  movel([0.496334, -1.374205, -2.584112, -0.754072, 1.570796, 2.067130],accel_mss,speed_ms,0,blend_radius_m)
  speed_ms = 0.05
  movel([0.496334, -1.321205, -2.558075, -0.833109, 1.570796, 2.067130],accel_mss,speed_ms,0,blend_radius_m)
  speed_ms = 0.051
  movel([0.496334, -1.311367, -2.552605, -0.848418, 1.570796, 2.067130],accel_mss,speed_ms,0,blend_radius_m)
  movel([0.393115, -1.332740, -2.538777, -0.840872, 1.570796, 1.963912],accel_mss,speed_ms,0,blend_radius_m)
  movel([0.393115, -1.362611, -2.554595, -0.795183, 1.570796, 1.963912],accel_mss,speed_ms,0,blend_radius_m)
  speed_ms = 0.017
  movel([0.393115, -1.394662, -2.569610, -0.748117, 1.570796, 1.963912],accel_mss,speed_ms,0,blend_radius_m)
  speed_ms = 0.051
  movel([0.404241, -1.368810, -2.587836, -0.755743, 1.570796, 1.975037],accel_mss,speed_ms,0,blend_radius_m)
  movel([0.405839, -1.365130, -2.590352, -0.756907, 1.570796, 1.976635],accel_mss,speed_ms,0,blend_radius_m)
  movel([0.405852, -1.365099, -2.590373, -0.756917, 1.570796, 1.976648],accel_mss,speed_ms,0,blend_radius_m)
  movel([0.406880, -1.363267, -2.591618, -0.757504, 1.570796, 1.977677],accel_mss,speed_ms,0,blend_radius_m)
  movel([0.408799, -1.360504, -2.593487, -0.758397, 1.570796, 1.979595],accel_mss,speed_ms,0,blend_radius_m)
  movel([0.410954, -1.358071, -2.595125, -0.759194, 1.570796, 1.981750],accel_mss,speed_ms,0,blend_radius_m)
  movel([0.413315, -1.355969, -2.596532, -0.759888, 1.570796, 1.984111],accel_mss,speed_ms,0,blend_radius_m)
  movel([0.415848, -1.354210, -2.597705, -0.760474, 1.570796, 1.986644],accel_mss,speed_ms,0,blend_radius_m)
  movel([0.418507, -1.352814, -2.598633, -0.760942, 1.570796, 1.989304],accel_mss,speed_ms,0,blend_radius_m)
  movel([0.421235, -1.351821, -2.599292, -0.761276, 1.570796, 1.992031],accel_mss,speed_ms,0,blend_radius_m)
  movel([0.423950, -1.351263, -2.599661, -0.761465, 1.570796, 1.994746],accel_mss,speed_ms,0,blend_radius_m)
  movel([0.426550, -1.351176, -2.599718, -0.761494, 1.570796, 1.997346],accel_mss,speed_ms,0,blend_radius_m)
  movel([0.428920, -1.351576, -2.599454, -0.761359, 1.570796, 1.999716],accel_mss,speed_ms,0,blend_radius_m)
  movel([0.430958, -1.352450, -2.598875, -0.761064, 1.570796, 2.001755],accel_mss,speed_ms,0,blend_radius_m)
  movel([0.432577, -1.353767, -2.598000, -0.760622, 1.570796, 2.003373],accel_mss,speed_ms,0,blend_radius_m)
  movel([0.433730, -1.355485, -2.596855, -0.760049, 1.570796, 2.004526],accel_mss,speed_ms,0,blend_radius_m)
  movel([0.434381, -1.357566, -2.595463, -0.759360, 1.570796, 2.005178],accel_mss,speed_ms,0,blend_radius_m)
  movel([0.434519, -1.359977, -2.593843, -0.758569, 1.570796, 2.005316],accel_mss,speed_ms,0,blend_radius_m)
  movel([0.434118, -1.362706, -2.591999, -0.757684, 1.570796, 2.004915],accel_mss,speed_ms,0,blend_radius_m)
  movel([0.433161, -1.365745, -2.589933, -0.756712, 1.570796, 2.003958],accel_mss,speed_ms,0,blend_radius_m)
  movel([0.431608, -1.369097, -2.587639, -0.755653, 1.570796, 2.002405],accel_mss,speed_ms,0,blend_radius_m)
  movel([0.430424, -1.371178, -2.586206, -0.755005, 1.570796, 2.001221],accel_mss,speed_ms,0,blend_radius_m)
  movel([0.439654, -1.371318, -2.586109, -0.754961, 1.570796, 2.010450],accel_mss,speed_ms,0,blend_radius_m)
  movel([0.436246, -1.378584, -2.581058, -0.752746, 1.570796, 2.007043],accel_mss,speed_ms,0,blend_radius_m)
  movel([0.410431, -1.378416, -2.581176, -0.752797, 1.570796, 1.981228],accel_mss,speed_ms,0,blend_radius_m)
  movel([0.413657, -1.371140, -2.586232, -0.755016, 1.570796, 1.984454],accel_mss,speed_ms,0,blend_radius_m)
  movel([0.422970, -1.371126, -2.586242, -0.755021, 1.570796, 1.993766],accel_mss,speed_ms,0,blend_radius_m)
  movel([0.424851, -1.367135, -2.588983, -0.756271, 1.570796, 1.995647],accel_mss,speed_ms,0,blend_radius_m)
  movel([0.425504, -1.365495, -2.590103, -0.756791, 1.570796, 1.996301],accel_mss,speed_ms,0,blend_radius_m)
  movel([0.425953, -1.364067, -2.591075, -0.757247, 1.570796, 1.996749],accel_mss,speed_ms,0,blend_radius_m)
  movel([0.426189, -1.362920, -2.591853, -0.757615, 1.570796, 1.996985],accel_mss,speed_ms,0,blend_radius_m)
  movel([0.426258, -1.361974, -2.592494, -0.757921, 1.570796, 1.997054],accel_mss,speed_ms,0,blend_radius_m)
  movel([0.426182, -1.361187, -2.593026, -0.758176, 1.570796, 1.996979],accel_mss,speed_ms,0,blend_radius_m)
  movel([0.425983, -1.360532, -2.593469, -0.758388, 1.570796, 1.996779],accel_mss,speed_ms,0,blend_radius_m)
  movel([0.425209, -1.359528, -2.594145, -0.758716, 1.570796, 1.996006],accel_mss,speed_ms,0,blend_radius_m)
  movel([0.423937, -1.358920, -2.594554, -0.758915, 1.570796, 1.994733],accel_mss,speed_ms,0,blend_radius_m)
  movel([0.422360, -1.358709, -2.594696, -0.758984, 1.570796, 1.993157],accel_mss,speed_ms,0,blend_radius_m)
  movel([0.421052, -1.358839, -2.594608, -0.758941, 1.570796, 1.991849],accel_mss,speed_ms,0,blend_radius_m)
  movel([0.419197, -1.359405, -2.594228, -0.758756, 1.570796, 1.989993],accel_mss,speed_ms,0,blend_radius_m)
  movel([0.417336, -1.360395, -2.593561, -0.758433, 1.570796, 1.988133],accel_mss,speed_ms,0,blend_radius_m)
  movel([0.415631, -1.361734, -2.592657, -0.757998, 1.570796, 1.986428],accel_mss,speed_ms,0,blend_radius_m)
  movel([0.414239, -1.363307, -2.591591, -0.757491, 1.570796, 1.985036],accel_mss,speed_ms,0,blend_radius_m)
  movel([0.413316, -1.364898, -2.590509, -0.756981, 1.570796, 1.984112],accel_mss,speed_ms,0,blend_radius_m)
  movel([0.402881, -1.388680, -2.573914, -0.749795, 1.570796, 1.973677],accel_mss,speed_ms,0,blend_radius_m)
  movel([0.400271, -1.389775, -2.573130, -0.749484, 1.570796, 1.971067],accel_mss,speed_ms,0,blend_radius_m)
  movel([0.397416, -1.391364, -2.571989, -0.749036, 1.570796, 1.968213],accel_mss,speed_ms,0,blend_radius_m)
  movel([0.394707, -1.393294, -2.570599, -0.748496, 1.570796, 1.965504],accel_mss,speed_ms,0,blend_radius_m)
  movel([0.393115, -1.394662, -2.569610, -0.748117, 1.570796, 1.963912],accel_mss,speed_ms,0,blend_radius_m)
  speed_ms = 0.05
  movel([0.393115, -1.342458, -2.544135, -0.825796, 1.570796, 1.963912],accel_mss,speed_ms,0,blend_radius_m)
  speed_ms = 0.051
  movel([0.393115, -1.332740, -2.538777, -0.840872, 1.570796, 1.963912],accel_mss,speed_ms,0,blend_radius_m)
  movel([0.435741, -1.287387, -2.567433, -0.857569, 1.570796, 2.006537],accel_mss,speed_ms,0,blend_radius_m)
  movel([0.435741, -1.318075, -2.583967, -0.810347, 1.570796, 2.006537],accel_mss,speed_ms,0,blend_radius_m)
  speed_ms = 0.017
  movel([0.435741, -1.351197, -2.599704, -0.761487, 1.570796, 2.006537],accel_mss,speed_ms,0,blend_radius_m)
  speed_ms = 0.051
  movel([0.437149, -1.352936, -2.598552, -0.760901, 1.570796, 2.007945],accel_mss,speed_ms,0,blend_radius_m)
  movel([0.438075, -1.355027, -2.597161, -0.760201, 1.570796, 2.008871],accel_mss,speed_ms,0,blend_radius_m)
  movel([0.438486, -1.357407, -2.595570, -0.759412, 1.570796, 2.009283],accel_mss,speed_ms,0,blend_radius_m)
  movel([0.438495, -1.358723, -2.594686, -0.758979, 1.570796, 2.009291],accel_mss,speed_ms,0,blend_radius_m)
  movel([0.462025, -1.359314, -2.594289, -0.758786, 1.570796, 2.032822],accel_mss,speed_ms,0,blend_radius_m)
  movel([0.462701, -1.359339, -2.594272, -0.758778, 1.570796, 2.033497],accel_mss,speed_ms,0,blend_radius_m)
  movel([0.464185, -1.359628, -2.594078, -0.758683, 1.570796, 2.034981],accel_mss,speed_ms,0,blend_radius_m)
  movel([0.465346, -1.360355, -2.593588, -0.758446, 1.570796, 2.036142],accel_mss,speed_ms,0,blend_radius_m)
  movel([0.466106, -1.361489, -2.592823, -0.758078, 1.570796, 2.036902],accel_mss,speed_ms,0,blend_radius_m)
  movel([0.466384, -1.362949, -2.591834, -0.757606, 1.570796, 2.037180],accel_mss,speed_ms,0,blend_radius_m)
  movel([0.466139, -1.364611, -2.590705, -0.757073, 1.570796, 2.036935],accel_mss,speed_ms,0,blend_radius_m)
  movel([0.465653, -1.365840, -2.589867, -0.756681, 1.570796, 2.036450],accel_mss,speed_ms,0,blend_radius_m)
  movel([0.464415, -1.367759, -2.588556, -0.756074, 1.570796, 2.035211],accel_mss,speed_ms,0,blend_radius_m)
  movel([0.463055, -1.369182, -2.587580, -0.755627, 1.570796, 2.033851],accel_mss,speed_ms,0,blend_radius_m)
  movel([0.461556, -1.370238, -2.586854, -0.755297, 1.570796, 2.032352],accel_mss,speed_ms,0,blend_radius_m)
  movel([0.459850, -1.371005, -2.586326, -0.755058, 1.570796, 2.030646],accel_mss,speed_ms,0,blend_radius_m)
  movel([0.457837, -1.371508, -2.585979, -0.754902, 1.570796, 2.028633],accel_mss,speed_ms,0,blend_radius_m)
  movel([0.455379, -1.371731, -2.585825, -0.754833, 1.570796, 2.026175],accel_mss,speed_ms,0,blend_radius_m)
  movel([0.452224, -1.371654, -2.585878, -0.754857, 1.570796, 2.023020],accel_mss,speed_ms,0,blend_radius_m)
  movel([0.450446, -1.371539, -2.585957, -0.754893, 1.570796, 2.021242],accel_mss,speed_ms,0,blend_radius_m)
  movel([0.454930, -1.362246, -2.592310, -0.757833, 1.570796, 2.025727],accel_mss,speed_ms,0,blend_radius_m)
  movel([0.447579, -1.362047, -2.592445, -0.757897, 1.570796, 2.018376],accel_mss,speed_ms,0,blend_radius_m)
  movel([0.435434, -1.387753, -2.574576, -0.750060, 1.570796, 2.006230],accel_mss,speed_ms,0,blend_radius_m)
  movel([0.442596, -1.387945, -2.574439, -0.750005, 1.570796, 2.013392],accel_mss,speed_ms,0,blend_radius_m)
  movel([0.446788, -1.379158, -2.580657, -0.752575, 1.570796, 2.017584],accel_mss,speed_ms,0,blend_radius_m)
  movel([0.446881, -1.378963, -2.580793, -0.752633, 1.570796, 2.017678],accel_mss,speed_ms,0,blend_radius_m)
  movel([0.446911, -1.378901, -2.580837, -0.752651, 1.570796, 2.017707],accel_mss,speed_ms,0,blend_radius_m)
  movel([0.450255, -1.379295, -2.580561, -0.752534, 1.570796, 2.021051],accel_mss,speed_ms,0,blend_radius_m)
  movel([0.453469, -1.379222, -2.580611, -0.752555, 1.570796, 2.024265],accel_mss,speed_ms,0,blend_radius_m)
  movel([0.456549, -1.378732, -2.580955, -0.752702, 1.570796, 2.027346],accel_mss,speed_ms,0,blend_radius_m)
  movel([0.459488, -1.377858, -2.581566, -0.752964, 1.570796, 2.030284],accel_mss,speed_ms,0,blend_radius_m)
  movel([0.462280, -1.376631, -2.582424, -0.753334, 1.570796, 2.033076],accel_mss,speed_ms,0,blend_radius_m)
  movel([0.464904, -1.375072, -2.583510, -0.753807, 1.570796, 2.035701],accel_mss,speed_ms,0,blend_radius_m)
  movel([0.467331, -1.373214, -2.584799, -0.754376, 1.570796, 2.038128],accel_mss,speed_ms,0,blend_radius_m)
  movel([0.469519, -1.371083, -2.586272, -0.755034, 1.570796, 2.040315],accel_mss,speed_ms,0,blend_radius_m)
  movel([0.471402, -1.368739, -2.587884, -0.755766, 1.570796, 2.042198],accel_mss,speed_ms,0,blend_radius_m)
  movel([0.472907, -1.366256, -2.589584, -0.756549, 1.570796, 2.043703],accel_mss,speed_ms,0,blend_radius_m)
  movel([0.473966, -1.363730, -2.591304, -0.757355, 1.570796, 2.044762],accel_mss,speed_ms,0,blend_radius_m)
  movel([0.474528, -1.361267, -2.592972, -0.758150, 1.570796, 2.045324],accel_mss,speed_ms,0,blend_radius_m)
  movel([0.474563, -1.358966, -2.594523, -0.758900, 1.570796, 2.045359],accel_mss,speed_ms,0,blend_radius_m)
  movel([0.474065, -1.356904, -2.595906, -0.759578, 1.570796, 2.044861],accel_mss,speed_ms,0,blend_radius_m)
  movel([0.473042, -1.355135, -2.597089, -0.760165, 1.570796, 2.043838],accel_mss,speed_ms,0,blend_radius_m)
  movel([0.471495, -1.353700, -2.598045, -0.760644, 1.570796, 2.042292],accel_mss,speed_ms,0,blend_radius_m)
  movel([0.469420, -1.352631, -2.598755, -0.761004, 1.570796, 2.040217],accel_mss,speed_ms,0,blend_radius_m)
  movel([0.466801, -1.351958, -2.599201, -0.761230, 1.570796, 2.037597],accel_mss,speed_ms,0,blend_radius_m)
  movel([0.466254, -1.351881, -2.599252, -0.761256, 1.570796, 2.037050],accel_mss,speed_ms,0,blend_radius_m)
  movel([0.435741, -1.351197, -2.599704, -0.761487, 1.570796, 2.006537],accel_mss,speed_ms,0,blend_radius_m)
  speed_ms = 0.05
  movel([0.435741, -1.297350, -2.573030, -0.842009, 1.570796, 2.006537],accel_mss,speed_ms,0,blend_radius_m)
  speed_ms = 0.051
  movel([0.435741, -1.287387, -2.567433, -0.857569, 1.570796, 2.006537],accel_mss,speed_ms,0,blend_radius_m)
  movel([0.468006, -1.313184, -2.551452, -0.847754, 1.570796, 2.038802],accel_mss,speed_ms,0,blend_radius_m)
  movel([0.468006, -1.343421, -2.567577, -0.801391, 1.570796, 2.038802],accel_mss,speed_ms,0,blend_radius_m)
  speed_ms = 0.017
  movel([0.468006, -1.375946, -2.582901, -0.753542, 1.570796, 2.038802],accel_mss,speed_ms,0,blend_radius_m)
  speed_ms = 0.051
  movel([0.456016, -1.400133, -2.565628, -0.746628, 1.570796, 2.026813],accel_mss,speed_ms,0,blend_radius_m)
  movel([0.453789, -1.404662, -2.562298, -0.745429, 1.570796, 2.024585],accel_mss,speed_ms,0,blend_radius_m)
  movel([0.453641, -1.404968, -2.562072, -0.745349, 1.570796, 2.024437],accel_mss,speed_ms,0,blend_radius_m)
  movel([0.452579, -1.406671, -2.560812, -0.744907, 1.570796, 2.023375],accel_mss,speed_ms,0,blend_radius_m)
  movel([0.450661, -1.409191, -2.558938, -0.744260, 1.570796, 2.021458],accel_mss,speed_ms,0,blend_radius_m)
  movel([0.448563, -1.411364, -2.557315, -0.743710, 1.570796, 2.019359],accel_mss,speed_ms,0,blend_radius_m)
  movel([0.446304, -1.413204, -2.555935, -0.743250, 1.570796, 2.017100],accel_mss,speed_ms,0,blend_radius_m)
  movel([0.443919, -1.414710, -2.554802, -0.742877, 1.570796, 2.014715],accel_mss,speed_ms,0,blend_radius_m)
  movel([0.441440, -1.415871, -2.553926, -0.742592, 1.570796, 2.012236],accel_mss,speed_ms,0,blend_radius_m)
  movel([0.438915, -1.416664, -2.553326, -0.742399, 1.570796, 2.009711],accel_mss,speed_ms,0,blend_radius_m)
  movel([0.436416, -1.417065, -2.553023, -0.742301, 1.570796, 2.007212],accel_mss,speed_ms,0,blend_radius_m)
  movel([0.434024, -1.417050, -2.553035, -0.742305, 1.570796, 2.004820],accel_mss,speed_ms,0,blend_radius_m)
  movel([0.431843, -1.416611, -2.553367, -0.742411, 1.570796, 2.002639],accel_mss,speed_ms,0,blend_radius_m)
  movel([0.429962, -1.415757, -2.554012, -0.742620, 1.570796, 2.000758],accel_mss,speed_ms,0,blend_radius_m)
  movel([0.428455, -1.414516, -2.554948, -0.742925, 1.570796, 1.999251],accel_mss,speed_ms,0,blend_radius_m)
  movel([0.427374, -1.412916, -2.556151, -0.743322, 1.570796, 1.998171],accel_mss,speed_ms,0,blend_radius_m)
  movel([0.426747, -1.410989, -2.557595, -0.743804, 1.570796, 1.997543],accel_mss,speed_ms,0,blend_radius_m)
  movel([0.426600, -1.408754, -2.559264, -0.744372, 1.570796, 1.997396],accel_mss,speed_ms,0,blend_radius_m)
  movel([0.426957, -1.406212, -2.561152, -0.745025, 1.570796, 1.997753],accel_mss,speed_ms,0,blend_radius_m)
  movel([0.427853, -1.403363, -2.563256, -0.745769, 1.570796, 1.998650],accel_mss,speed_ms,0,blend_radius_m)
  movel([0.429335, -1.400194, -2.565584, -0.746612, 1.570796, 2.000131],accel_mss,speed_ms,0,blend_radius_m)
  movel([0.430468, -1.398225, -2.567022, -0.747142, 1.570796, 2.001264],accel_mss,speed_ms,0,blend_radius_m)
  movel([0.421486, -1.398069, -2.567136, -0.747184, 1.570796, 1.992282],accel_mss,speed_ms,0,blend_radius_m)
  movel([0.424715, -1.391019, -2.572237, -0.749133, 1.570796, 1.995511],accel_mss,speed_ms,0,blend_radius_m)
  movel([0.449964, -1.391682, -2.571760, -0.748946, 1.570796, 2.020760],accel_mss,speed_ms,0,blend_radius_m)
  movel([0.446570, -1.398709, -2.566669, -0.747011, 1.570796, 2.017367],accel_mss,speed_ms,0,blend_radius_m)
  movel([0.437657, -1.398406, -2.566890, -0.747093, 1.570796, 2.008453],accel_mss,speed_ms,0,blend_radius_m)
  movel([0.435797, -1.402197, -2.564115, -0.746078, 1.570796, 2.006593],accel_mss,speed_ms,0,blend_radius_m)
  movel([0.435154, -1.403745, -2.562975, -0.745669, 1.570796, 2.005951],accel_mss,speed_ms,0,blend_radius_m)
  movel([0.434713, -1.405089, -2.561983, -0.745317, 1.570796, 2.005509],accel_mss,speed_ms,0,blend_radius_m)
  movel([0.434481, -1.406166, -2.561185, -0.745037, 1.570796, 2.005277],accel_mss,speed_ms,0,blend_radius_m)
  movel([0.434406, -1.407058, -2.560524, -0.744807, 1.570796, 2.005202],accel_mss,speed_ms,0,blend_radius_m)
  movel([0.434470, -1.407800, -2.559974, -0.744616, 1.570796, 2.005266],accel_mss,speed_ms,0,blend_radius_m)
  movel([0.434651, -1.408420, -2.559512, -0.744457, 1.570796, 2.005447],accel_mss,speed_ms,0,blend_radius_m)
  movel([0.435365, -1.409380, -2.558797, -0.744212, 1.570796, 2.006161],accel_mss,speed_ms,0,blend_radius_m)
  movel([0.436549, -1.409986, -2.558345, -0.744058, 1.570796, 2.007345],accel_mss,speed_ms,0,blend_radius_m)
  movel([0.438023, -1.410235, -2.558159, -0.743995, 1.570796, 2.008819],accel_mss,speed_ms,0,blend_radius_m)
  movel([0.439241, -1.410163, -2.558213, -0.744013, 1.570796, 2.010038],accel_mss,speed_ms,0,blend_radius_m)
  movel([0.440983, -1.409705, -2.558554, -0.744129, 1.570796, 2.011779],accel_mss,speed_ms,0,blend_radius_m)
  movel([0.442739, -1.408855, -2.559189, -0.744346, 1.570796, 2.013535],accel_mss,speed_ms,0,blend_radius_m)
  movel([0.444367, -1.407667, -2.560072, -0.744650, 1.570796, 2.015163],accel_mss,speed_ms,0,blend_radius_m)
  movel([0.445716, -1.406238, -2.561132, -0.745018, 1.570796, 2.016512],accel_mss,speed_ms,0,blend_radius_m)
  movel([0.446637, -1.404764, -2.562223, -0.745402, 1.570796, 2.017433],accel_mss,speed_ms,0,blend_radius_m)
  movel([0.457925, -1.381620, -2.578926, -0.751843, 1.570796, 2.028721],accel_mss,speed_ms,0,blend_radius_m)
  movel([0.460558, -1.380630, -2.579623, -0.752136, 1.570796, 2.031354],accel_mss,speed_ms,0,blend_radius_m)
  movel([0.463484, -1.379143, -2.580667, -0.752579, 1.570796, 2.034281],accel_mss,speed_ms,0,blend_radius_m)
  movel([0.466307, -1.377290, -2.581964, -0.753135, 1.570796, 2.037103],accel_mss,speed_ms,0,blend_radius_m)
  movel([0.468006, -1.375946, -2.582901, -0.753542, 1.570796, 2.038802],accel_mss,speed_ms,0,blend_radius_m)
  speed_ms = 0.05
  movel([0.468006, -1.323012, -2.556913, -0.832464, 1.570796, 2.038802],accel_mss,speed_ms,0,blend_radius_m)
  speed_ms = 0.051
  movel([0.468006, -1.313184, -2.551452, -0.847754, 1.570796, 2.038802],accel_mss,speed_ms,0,blend_radius_m)
  movel([0.425547, -1.355903, -2.523122, -0.833364, 1.570796, 1.996343],accel_mss,speed_ms,0,blend_radius_m)
  movel([0.425547, -1.385315, -2.538580, -0.788493, 1.570796, 1.996343],accel_mss,speed_ms,0,blend_radius_m)
  speed_ms = 0.017
  movel([0.425547, -1.416785, -2.553235, -0.742369, 1.570796, 1.996343],accel_mss,speed_ms,0,blend_radius_m)
  speed_ms = 0.051
  movel([0.403473, -1.416474, -2.553470, -0.742445, 1.570796, 1.974270],accel_mss,speed_ms,0,blend_radius_m)
  movel([0.396842, -1.416472, -2.553471, -0.742445, 1.570796, 1.967639],accel_mss,speed_ms,0,blend_radius_m)
  movel([0.396831, -1.416472, -2.553471, -0.742445, 1.570796, 1.967627],accel_mss,speed_ms,0,blend_radius_m)
  movel([0.395180, -1.416267, -2.553626, -0.742495, 1.570796, 1.965977],accel_mss,speed_ms,0,blend_radius_m)
  movel([0.392846, -1.415632, -2.554106, -0.742651, 1.570796, 1.963642],accel_mss,speed_ms,0,blend_radius_m)
  movel([0.390981, -1.414656, -2.554843, -0.742891, 1.570796, 1.961777],accel_mss,speed_ms,0,blend_radius_m)
  movel([0.389571, -1.413365, -2.555814, -0.743210, 1.570796, 1.960368],accel_mss,speed_ms,0,blend_radius_m)
  movel([0.388609, -1.411785, -2.557000, -0.743604, 1.570796, 1.959406],accel_mss,speed_ms,0,blend_radius_m)
  movel([0.388105, -1.409938, -2.558381, -0.744070, 1.570796, 1.958902],accel_mss,speed_ms,0,blend_radius_m)
  movel([0.388072, -1.407859, -2.559929, -0.744600, 1.570796, 1.958868],accel_mss,speed_ms,0,blend_radius_m)
  movel([0.388518, -1.405604, -2.561602, -0.745183, 1.570796, 1.959314],accel_mss,speed_ms,0,blend_radius_m)
  movel([0.389446, -1.403245, -2.563343, -0.745801, 1.570796, 1.960243],accel_mss,speed_ms,0,blend_radius_m)
  movel([0.390831, -1.400879, -2.565081, -0.746428, 1.570796, 1.961628],accel_mss,speed_ms,0,blend_radius_m)
  movel([0.392628, -1.398602, -2.566747, -0.747040, 1.570796, 1.963425],accel_mss,speed_ms,0,blend_radius_m)
  movel([0.394772, -1.396508, -2.568271, -0.747609, 1.570796, 1.965569],accel_mss,speed_ms,0,blend_radius_m)
  movel([0.397198, -1.394665, -2.569608, -0.748116, 1.570796, 1.967995],accel_mss,speed_ms,0,blend_radius_m)
  movel([0.399853, -1.393125, -2.570721, -0.748543, 1.570796, 1.970650],accel_mss,speed_ms,0,blend_radius_m)
  movel([0.402697, -1.391919, -2.571590, -0.748880, 1.570796, 1.973493],accel_mss,speed_ms,0,blend_radius_m)
  movel([0.405704, -1.391081, -2.572193, -0.749115, 1.570796, 1.976501],accel_mss,speed_ms,0,blend_radius_m)
  movel([0.408860, -1.390644, -2.572506, -0.749238, 1.570796, 1.979657],accel_mss,speed_ms,0,blend_radius_m)
  movel([0.412150, -1.390646, -2.572505, -0.749238, 1.570796, 1.982946],accel_mss,speed_ms,0,blend_radius_m)
  movel([0.414108, -1.390866, -2.572347, -0.749176, 1.570796, 1.984905],accel_mss,speed_ms,0,blend_radius_m)
  movel([0.418149, -1.381867, -2.578751, -0.751770, 1.570796, 1.988945],accel_mss,speed_ms,0,blend_radius_m)
  movel([0.425423, -1.381914, -2.578718, -0.751757, 1.570796, 1.996219],accel_mss,speed_ms,0,blend_radius_m)
  movel([0.414112, -1.406828, -2.560695, -0.744866, 1.570796, 1.984908],accel_mss,speed_ms,0,blend_radius_m)
  movel([0.407010, -1.406787, -2.560726, -0.744877, 1.570796, 1.977806],accel_mss,speed_ms,0,blend_radius_m)
  movel([0.410920, -1.398011, -2.567178, -0.747200, 1.570796, 1.981717],accel_mss,speed_ms,0,blend_radius_m)
  movel([0.407049, -1.397939, -2.567230, -0.747220, 1.570796, 1.977845],accel_mss,speed_ms,0,blend_radius_m)
  movel([0.405413, -1.398026, -2.567167, -0.747196, 1.570796, 1.976209],accel_mss,speed_ms,0,blend_radius_m)
  movel([0.403942, -1.398220, -2.567026, -0.747143, 1.570796, 1.974739],accel_mss,speed_ms,0,blend_radius_m)
  movel([0.402713, -1.398494, -2.566826, -0.747069, 1.570796, 1.973509],accel_mss,speed_ms,0,blend_radius_m)
  movel([0.401648, -1.398841, -2.566572, -0.746975, 1.570796, 1.972444],accel_mss,speed_ms,0,blend_radius_m)
  movel([0.400712, -1.399250, -2.566274, -0.746865, 1.570796, 1.971508],accel_mss,speed_ms,0,blend_radius_m)
  movel([0.399874, -1.399720, -2.565930, -0.746739, 1.570796, 1.970671],accel_mss,speed_ms,0,blend_radius_m)
  movel([0.398410, -1.400878, -2.565082, -0.746428, 1.570796, 1.969206],accel_mss,speed_ms,0,blend_radius_m)
  movel([0.397202, -1.402325, -2.564020, -0.746044, 1.570796, 1.967999],accel_mss,speed_ms,0,blend_radius_m)
  movel([0.396320, -1.403889, -2.562869, -0.745631, 1.570796, 1.967117],accel_mss,speed_ms,0,blend_radius_m)
  movel([0.395938, -1.405045, -2.562015, -0.745329, 1.570796, 1.966735],accel_mss,speed_ms,0,blend_radius_m)
  movel([0.395831, -1.406526, -2.560919, -0.744944, 1.570796, 1.966627],accel_mss,speed_ms,0,blend_radius_m)
  movel([0.396199, -1.407832, -2.559950, -0.744608, 1.570796, 1.966995],accel_mss,speed_ms,0,blend_radius_m)
  movel([0.397028, -1.408849, -2.559193, -0.744347, 1.570796, 1.967824],accel_mss,speed_ms,0,blend_radius_m)
  movel([0.398251, -1.409481, -2.558722, -0.744186, 1.570796, 1.969048],accel_mss,speed_ms,0,blend_radius_m)
  movel([0.399687, -1.409681, -2.558573, -0.744135, 1.570796, 1.970483],accel_mss,speed_ms,0,blend_radius_m)
  movel([0.422863, -1.409863, -2.558437, -0.744089, 1.570796, 1.993659],accel_mss,speed_ms,0,blend_radius_m)
  movel([0.422993, -1.411906, -2.556909, -0.743574, 1.570796, 1.993789],accel_mss,speed_ms,0,blend_radius_m)
  movel([0.423592, -1.413991, -2.555343, -0.743055, 1.570796, 1.994388],accel_mss,speed_ms,0,blend_radius_m)
  movel([0.424651, -1.415802, -2.553978, -0.742609, 1.570796, 1.995448],accel_mss,speed_ms,0,blend_radius_m)
  movel([0.425547, -1.416785, -2.553235, -0.742369, 1.570796, 1.996343],accel_mss,speed_ms,0,blend_radius_m)
  speed_ms = 0.05
  movel([0.425547, -1.365481, -2.528361, -0.818547, 1.570796, 1.996343],accel_mss,speed_ms,0,blend_radius_m)
  speed_ms = 0.051
  movel([0.425547, -1.355903, -2.523122, -0.833364, 1.570796, 1.996343],accel_mss,speed_ms,0,blend_radius_m)
  movel([0.496386, -1.351291, -2.526295, -0.834803, 1.570796, 2.067183],accel_mss,speed_ms,0,blend_radius_m)
  movel([0.496386, -1.380797, -2.541825, -0.789767, 1.570796, 2.067183],accel_mss,speed_ms,0,blend_radius_m)
  speed_ms = 0.017
  movel([0.496386, -1.412384, -2.556551, -0.743454, 1.570796, 2.067183],accel_mss,speed_ms,0,blend_radius_m)
  speed_ms = 0.051
  movel([0.494250, -1.412916, -2.556152, -0.743322, 1.570796, 2.065047],accel_mss,speed_ms,0,blend_radius_m)
  movel([0.492155, -1.413824, -2.555469, -0.743096, 1.570796, 2.062951],accel_mss,speed_ms,0,blend_radius_m)
  movel([0.490635, -1.414706, -2.554805, -0.742878, 1.570796, 2.061431],accel_mss,speed_ms,0,blend_radius_m)
  movel([0.498563, -1.433670, -2.540242, -0.738476, 1.570796, 2.069360],accel_mss,speed_ms,0,blend_radius_m)
  movel([0.507323, -1.428619, -2.544174, -0.739595, 1.570796, 2.078119],accel_mss,speed_ms,0,blend_radius_m)
  movel([0.504979, -1.429334, -2.543621, -0.739435, 1.570796, 2.075776],accel_mss,speed_ms,0,blend_radius_m)
  movel([0.502994, -1.429562, -2.543443, -0.739383, 1.570796, 2.073791],accel_mss,speed_ms,0,blend_radius_m)
  movel([0.501213, -1.429380, -2.543585, -0.739424, 1.570796, 2.072009],accel_mss,speed_ms,0,blend_radius_m)
  movel([0.499589, -1.428783, -2.544047, -0.739558, 1.570796, 2.070385],accel_mss,speed_ms,0,blend_radius_m)
  movel([0.498113, -1.427739, -2.544855, -0.739794, 1.570796, 2.068909],accel_mss,speed_ms,0,blend_radius_m)
  movel([0.496789, -1.426184, -2.546056, -0.740149, 1.570796, 2.067585],accel_mss,speed_ms,0,blend_radius_m)
  movel([0.495653, -1.424054, -2.547695, -0.740640, 1.570796, 2.066450],accel_mss,speed_ms,0,blend_radius_m)
  movel([0.495357, -1.423295, -2.548277, -0.740817, 1.570796, 2.066154],accel_mss,speed_ms,0,blend_radius_m)
  movel([0.496802, -1.422585, -2.548821, -0.740983, 1.570796, 2.067599],accel_mss,speed_ms,0,blend_radius_m)
  movel([0.498935, -1.421858, -2.549377, -0.741154, 1.570796, 2.069732],accel_mss,speed_ms,0,blend_radius_m)
  movel([0.501190, -1.421465, -2.549677, -0.741247, 1.570796, 2.071986],accel_mss,speed_ms,0,blend_radius_m)
  movel([0.503721, -1.421404, -2.549724, -0.741261, 1.570796, 2.074517],accel_mss,speed_ms,0,blend_radius_m)
  movel([0.506892, -1.421700, -2.549497, -0.741191, 1.570796, 2.077688],accel_mss,speed_ms,0,blend_radius_m)
  movel([0.508953, -1.421976, -2.549287, -0.741126, 1.570796, 2.079749],accel_mss,speed_ms,0,blend_radius_m)
  movel([0.511017, -1.422212, -2.549106, -0.741071, 1.570796, 2.081813],accel_mss,speed_ms,0,blend_radius_m)
  movel([0.512879, -1.422311, -2.549031, -0.741048, 1.570796, 2.083675],accel_mss,speed_ms,0,blend_radius_m)
  movel([0.514361, -1.422273, -2.549060, -0.741057, 1.570796, 2.085157],accel_mss,speed_ms,0,blend_radius_m)
  movel([0.516717, -1.421930, -2.549322, -0.741137, 1.570796, 2.087514],accel_mss,speed_ms,0,blend_radius_m)
  movel([0.519106, -1.421259, -2.549835, -0.741296, 1.570796, 2.089902],accel_mss,speed_ms,0,blend_radius_m)
  movel([0.521253, -1.420298, -2.550567, -0.741524, 1.570796, 2.092049],accel_mss,speed_ms,0,blend_radius_m)
  movel([0.523071, -1.419109, -2.551472, -0.741808, 1.570796, 2.093867],accel_mss,speed_ms,0,blend_radius_m)
  movel([0.524605, -1.417699, -2.552542, -0.742147, 1.570796, 2.095402],accel_mss,speed_ms,0,blend_radius_m)
  movel([0.525885, -1.416058, -2.553785, -0.742546, 1.570796, 2.096681],accel_mss,speed_ms,0,blend_radius_m)
  movel([0.526903, -1.414161, -2.555215, -0.743013, 1.570796, 2.097699],accel_mss,speed_ms,0,blend_radius_m)
  movel([0.527617, -1.412010, -2.556831, -0.743548, 1.570796, 2.098413],accel_mss,speed_ms,0,blend_radius_m)
  movel([0.527962, -1.409636, -2.558606, -0.744147, 1.570796, 2.098758],accel_mss,speed_ms,0,blend_radius_m)
  movel([0.527865, -1.407145, -2.560460, -0.744784, 1.570796, 2.098662],accel_mss,speed_ms,0,blend_radius_m)
  movel([0.527282, -1.404723, -2.562253, -0.745413, 1.570796, 2.098079],accel_mss,speed_ms,0,blend_radius_m)
  movel([0.526229, -1.402597, -2.563820, -0.745972, 1.570796, 2.097026],accel_mss,speed_ms,0,blend_radius_m)
  movel([0.524809, -1.400967, -2.565017, -0.746405, 1.570796, 2.095605],accel_mss,speed_ms,0,blend_radius_m)
  movel([0.523535, -1.400104, -2.565650, -0.746636, 1.570796, 2.094332],accel_mss,speed_ms,0,blend_radius_m)
  movel([0.522574, -1.399712, -2.565936, -0.746741, 1.570796, 2.093370],accel_mss,speed_ms,0,blend_radius_m)
  movel([0.521144, -1.399562, -2.566046, -0.746781, 1.570796, 2.091941],accel_mss,speed_ms,0,blend_radius_m)
  movel([0.519713, -1.399841, -2.565842, -0.746706, 1.570796, 2.090509],accel_mss,speed_ms,0,blend_radius_m)
  movel([0.518321, -1.400499, -2.565360, -0.746530, 1.570796, 2.089117],accel_mss,speed_ms,0,blend_radius_m)
  movel([0.517042, -1.401495, -2.564630, -0.746264, 1.570796, 2.087839],accel_mss,speed_ms,0,blend_radius_m)
  movel([0.516004, -1.402743, -2.563713, -0.745933, 1.570796, 2.086801],accel_mss,speed_ms,0,blend_radius_m)
  movel([0.515361, -1.404091, -2.562720, -0.745578, 1.570796, 2.086157],accel_mss,speed_ms,0,blend_radius_m)
  movel([0.515210, -1.405299, -2.561828, -0.745262, 1.570796, 2.086007],accel_mss,speed_ms,0,blend_radius_m)
  movel([0.515554, -1.406380, -2.561027, -0.744982, 1.570796, 2.086350],accel_mss,speed_ms,0,blend_radius_m)
  movel([0.516416, -1.407204, -2.560416, -0.744769, 1.570796, 2.087212],accel_mss,speed_ms,0,blend_radius_m)
  movel([0.517279, -1.407592, -2.560128, -0.744669, 1.570796, 2.088075],accel_mss,speed_ms,0,blend_radius_m)
  movel([0.518096, -1.407710, -2.560040, -0.744639, 1.570796, 2.088893],accel_mss,speed_ms,0,blend_radius_m)
  movel([0.519202, -1.407488, -2.560205, -0.744696, 1.570796, 2.089998],accel_mss,speed_ms,0,blend_radius_m)
  movel([0.520433, -1.406863, -2.560669, -0.744857, 1.570796, 2.091230],accel_mss,speed_ms,0,blend_radius_m)
  movel([0.521857, -1.405770, -2.561479, -0.745140, 1.570796, 2.092653],accel_mss,speed_ms,0,blend_radius_m)
  movel([0.523464, -1.404168, -2.562663, -0.745558, 1.570796, 2.094260],accel_mss,speed_ms,0,blend_radius_m)
  movel([0.523573, -1.404048, -2.562751, -0.745589, 1.570796, 2.094369],accel_mss,speed_ms,0,blend_radius_m)
  movel([0.524385, -1.403902, -2.562859, -0.745628, 1.570796, 2.095181],accel_mss,speed_ms,0,blend_radius_m)
  movel([0.525389, -1.404028, -2.562766, -0.745595, 1.570796, 2.096185],accel_mss,speed_ms,0,blend_radius_m)
  movel([0.526064, -1.404552, -2.562380, -0.745458, 1.570796, 2.096860],accel_mss,speed_ms,0,blend_radius_m)
  movel([0.526402, -1.405475, -2.561697, -0.745217, 1.570796, 2.097199],accel_mss,speed_ms,0,blend_radius_m)
  movel([0.526323, -1.406784, -2.560727, -0.744877, 1.570796, 2.097119],accel_mss,speed_ms,0,blend_radius_m)
  movel([0.525762, -1.408332, -2.559577, -0.744479, 1.570796, 2.096558],accel_mss,speed_ms,0,blend_radius_m)
  movel([0.524768, -1.409827, -2.558464, -0.744098, 1.570796, 2.095564],accel_mss,speed_ms,0,blend_radius_m)
  movel([0.524179, -1.410451, -2.557998, -0.743940, 1.570796, 2.094975],accel_mss,speed_ms,0,blend_radius_m)
  movel([0.523546, -1.410986, -2.557598, -0.743805, 1.570796, 2.094342],accel_mss,speed_ms,0,blend_radius_m)
  movel([0.522160, -1.411793, -2.556994, -0.743602, 1.570796, 2.092957],accel_mss,speed_ms,0,blend_radius_m)
  movel([0.522122, -1.411809, -2.556982, -0.743598, 1.570796, 2.092918],accel_mss,speed_ms,0,blend_radius_m)
  movel([0.520402, -1.412510, -2.556456, -0.743423, 1.570796, 2.091198],accel_mss,speed_ms,0,blend_radius_m)
  movel([0.518013, -1.413155, -2.555972, -0.743262, 1.570796, 2.088809],accel_mss,speed_ms,0,blend_radius_m)
  movel([0.515460, -1.413467, -2.555737, -0.743185, 1.570796, 2.086257],accel_mss,speed_ms,0,blend_radius_m)
  movel([0.512586, -1.413441, -2.555757, -0.743191, 1.570796, 2.083382],accel_mss,speed_ms,0,blend_radius_m)
  movel([0.509044, -1.413037, -2.556060, -0.743292, 1.570796, 2.079841],accel_mss,speed_ms,0,blend_radius_m)
  movel([0.506535, -1.412642, -2.556357, -0.743390, 1.570796, 2.077331],accel_mss,speed_ms,0,blend_radius_m)
  movel([0.504024, -1.412280, -2.556629, -0.743481, 1.570796, 2.074820],accel_mss,speed_ms,0,blend_radius_m)
  movel([0.501612, -1.412053, -2.556799, -0.743537, 1.570796, 2.072409],accel_mss,speed_ms,0,blend_radius_m)
  movel([0.499823, -1.412015, -2.556827, -0.743547, 1.570796, 2.070619],accel_mss,speed_ms,0,blend_radius_m)
  movel([0.498273, -1.412102, -2.556762, -0.743525, 1.570796, 2.069069],accel_mss,speed_ms,0,blend_radius_m)
  movel([0.496386, -1.412384, -2.556551, -0.743454, 1.570796, 2.067183],accel_mss,speed_ms,0,blend_radius_m)
  speed_ms = 0.05
  movel([0.496386, -1.360898, -2.531558, -0.819933, 1.570796, 2.067183],accel_mss,speed_ms,0,blend_radius_m)
  speed_ms = 0.051
  movel([0.496386, -1.351291, -2.526295, -0.834803, 1.570796, 2.067183],accel_mss,speed_ms,0,blend_radius_m)
  movel([0.501294, -1.380106, -2.506003, -0.826280, 1.570796, 2.072091],accel_mss,speed_ms,0,blend_radius_m)
  movel([0.501294, -1.409013, -2.521091, -0.782286, 1.570796, 2.072091],accel_mss,speed_ms,0,blend_radius_m)
  speed_ms = 0.017
  movel([0.501294, -1.439855, -2.535375, -0.737159, 1.570796, 2.072091],accel_mss,speed_ms,0,blend_radius_m)
  speed_ms = 0.051
  movel([0.501364, -1.438344, -2.536570, -0.737475, 1.570796, 2.072160],accel_mss,speed_ms,0,blend_radius_m)
  movel([0.501902, -1.436575, -2.537964, -0.737850, 1.570796, 2.072698],accel_mss,speed_ms,0,blend_radius_m)
  movel([0.502852, -1.434869, -2.539304, -0.738216, 1.570796, 2.073649],accel_mss,speed_ms,0,blend_radius_m)
  movel([0.503411, -1.434165, -2.539855, -0.738369, 1.570796, 2.074207],accel_mss,speed_ms,0,blend_radius_m)
  movel([0.503999, -1.433568, -2.540323, -0.738498, 1.570796, 2.074796],accel_mss,speed_ms,0,blend_radius_m)
  movel([0.504606, -1.433084, -2.540701, -0.738604, 1.570796, 2.075402],accel_mss,speed_ms,0,blend_radius_m)
  movel([0.505876, -1.432412, -2.541226, -0.738751, 1.570796, 2.076673],accel_mss,speed_ms,0,blend_radius_m)
  movel([0.507182, -1.432148, -2.541432, -0.738809, 1.570796, 2.077978],accel_mss,speed_ms,0,blend_radius_m)
  movel([0.508066, -1.432194, -2.541395, -0.738799, 1.570796, 2.078863],accel_mss,speed_ms,0,blend_radius_m)
  movel([0.509244, -1.432844, -2.540888, -0.738657, 1.570796, 2.080041],accel_mss,speed_ms,0,blend_radius_m)
  movel([0.509920, -1.433743, -2.540185, -0.738460, 1.570796, 2.080716],accel_mss,speed_ms,0,blend_radius_m)
  movel([0.510117, -1.434828, -2.539336, -0.738225, 1.570796, 2.080914],accel_mss,speed_ms,0,blend_radius_m)
  movel([0.509853, -1.436017, -2.538403, -0.737969, 1.570796, 2.080649],accel_mss,speed_ms,0,blend_radius_m)
  movel([0.509157, -1.437210, -2.537464, -0.737715, 1.570796, 2.079953],accel_mss,speed_ms,0,blend_radius_m)
  movel([0.508088, -1.438286, -2.536615, -0.737487, 1.570796, 2.078884],accel_mss,speed_ms,0,blend_radius_m)
  movel([0.506729, -1.439143, -2.535939, -0.737307, 1.570796, 2.077525],accel_mss,speed_ms,0,blend_radius_m)
  movel([0.505151, -1.439703, -2.535495, -0.737190, 1.570796, 2.075947],accel_mss,speed_ms,0,blend_radius_m)
  movel([0.503715, -1.439905, -2.535335, -0.737148, 1.570796, 2.074511],accel_mss,speed_ms,0,blend_radius_m)
  movel([0.502898, -1.440772, -2.534649, -0.736968, 1.570796, 2.073694],accel_mss,speed_ms,0,blend_radius_m)
  movel([0.502527, -1.441638, -2.533961, -0.736790, 1.570796, 2.073324],accel_mss,speed_ms,0,blend_radius_m)
  movel([0.502557, -1.442533, -2.533250, -0.736607, 1.570796, 2.073353],accel_mss,speed_ms,0,blend_radius_m)
  movel([0.503041, -1.443448, -2.532520, -0.736420, 1.570796, 2.073837],accel_mss,speed_ms,0,blend_radius_m)
  movel([0.504021, -1.444249, -2.531882, -0.736258, 1.570796, 2.074818],accel_mss,speed_ms,0,blend_radius_m)
  movel([0.505332, -1.444698, -2.531523, -0.736168, 1.570796, 2.076129],accel_mss,speed_ms,0,blend_radius_m)
  movel([0.505913, -1.444738, -2.531491, -0.736160, 1.570796, 2.076710],accel_mss,speed_ms,0,blend_radius_m)
  movel([0.506013, -1.444735, -2.531493, -0.736161, 1.570796, 2.076810],accel_mss,speed_ms,0,blend_radius_m)
  movel([0.508325, -1.444424, -2.531742, -0.736223, 1.570796, 2.079121],accel_mss,speed_ms,0,blend_radius_m)
  movel([0.510402, -1.443778, -2.532257, -0.736353, 1.570796, 2.081199],accel_mss,speed_ms,0,blend_radius_m)
  movel([0.512273, -1.442835, -2.533009, -0.736545, 1.570796, 2.083070],accel_mss,speed_ms,0,blend_radius_m)
  movel([0.513958, -1.441610, -2.533984, -0.736796, 1.570796, 2.084755],accel_mss,speed_ms,0,blend_radius_m)
  movel([0.515462, -1.440103, -2.535179, -0.737107, 1.570796, 2.086259],accel_mss,speed_ms,0,blend_radius_m)
  movel([0.516762, -1.438317, -2.536591, -0.737481, 1.570796, 2.087558],accel_mss,speed_ms,0,blend_radius_m)
  movel([0.517807, -1.436265, -2.538208, -0.737916, 1.570796, 2.088604],accel_mss,speed_ms,0,blend_radius_m)
  movel([0.518520, -1.434013, -2.539974, -0.738402, 1.570796, 2.089316],accel_mss,speed_ms,0,blend_radius_m)
  movel([0.518819, -1.431676, -2.541800, -0.738913, 1.570796, 2.089615],accel_mss,speed_ms,0,blend_radius_m)
  movel([0.518653, -1.429447, -2.543533, -0.739409, 1.570796, 2.089450],accel_mss,speed_ms,0,blend_radius_m)
  movel([0.518009, -1.427400, -2.545118, -0.739871, 1.570796, 2.088805],accel_mss,speed_ms,0,blend_radius_m)
  movel([0.517775, -1.426940, -2.545473, -0.739976, 1.570796, 2.088572],accel_mss,speed_ms,0,blend_radius_m)
  movel([0.531403, -1.419285, -2.551338, -0.741765, 1.570796, 2.102199],accel_mss,speed_ms,0,blend_radius_m)
  movel([0.536550, -1.433923, -2.540045, -0.738421, 1.570796, 2.107347],accel_mss,speed_ms,0,blend_radius_m)
  movel([0.528022, -1.438600, -2.536368, -0.737421, 1.570796, 2.098818],accel_mss,speed_ms,0,blend_radius_m)
  movel([0.527776, -1.438735, -2.536261, -0.737393, 1.570796, 2.098573],accel_mss,speed_ms,0,blend_radius_m)
  movel([0.529435, -1.437274, -2.537414, -0.737702, 1.570796, 2.100232],accel_mss,speed_ms,0,blend_radius_m)
  movel([0.530798, -1.435628, -2.538708, -0.738053, 1.570796, 2.101594],accel_mss,speed_ms,0,blend_radius_m)
  movel([0.531867, -1.433791, -2.540148, -0.738450, 1.570796, 2.102664],accel_mss,speed_ms,0,blend_radius_m)
  movel([0.532619, -1.431766, -2.541730, -0.738894, 1.570796, 2.103415],accel_mss,speed_ms,0,blend_radius_m)
  movel([0.532999, -1.429585, -2.543425, -0.739378, 1.570796, 2.103795],accel_mss,speed_ms,0,blend_radius_m)
  movel([0.532952, -1.427341, -2.545163, -0.739885, 1.570796, 2.103748],accel_mss,speed_ms,0,blend_radius_m)
  movel([0.532435, -1.425198, -2.546816, -0.740376, 1.570796, 2.103231],accel_mss,speed_ms,0,blend_radius_m)
  movel([0.532418, -1.425154, -2.546849, -0.740386, 1.570796, 2.103214],accel_mss,speed_ms,0,blend_radius_m)
  movel([0.522682, -1.430574, -2.542657, -0.739158, 1.570796, 2.093478],accel_mss,speed_ms,0,blend_radius_m)
  movel([0.522463, -1.430698, -2.542561, -0.739130, 1.570796, 2.093259],accel_mss,speed_ms,0,blend_radius_m)
  movel([0.522402, -1.430731, -2.542535, -0.739123, 1.570796, 2.093198],accel_mss,speed_ms,0,blend_radius_m)
  movel([0.523214, -1.433581, -2.540313, -0.738496, 1.570796, 2.094010],accel_mss,speed_ms,0,blend_radius_m)
  movel([0.523471, -1.436241, -2.538226, -0.737921, 1.570796, 2.094267],accel_mss,speed_ms,0,blend_radius_m)
  movel([0.523250, -1.438696, -2.536291, -0.737401, 1.570796, 2.094046],accel_mss,speed_ms,0,blend_radius_m)
  movel([0.522620, -1.440937, -2.534518, -0.736934, 1.570796, 2.093417],accel_mss,speed_ms,0,blend_radius_m)
  movel([0.521637, -1.442957, -2.532912, -0.736520, 1.570796, 2.092433],accel_mss,speed_ms,0,blend_radius_m)
  movel([0.520354, -1.444747, -2.531483, -0.736158, 1.570796, 2.091150],accel_mss,speed_ms,0,blend_radius_m)
  movel([0.518812, -1.446300, -2.530240, -0.735848, 1.570796, 2.089609],accel_mss,speed_ms,0,blend_radius_m)
  movel([0.517050, -1.447597, -2.529200, -0.735592, 1.570796, 2.087847],accel_mss,speed_ms,0,blend_radius_m)
  movel([0.515113, -1.448608, -2.528386, -0.735395, 1.570796, 2.085909],accel_mss,speed_ms,0,blend_radius_m)
  movel([0.513057, -1.449295, -2.527833, -0.735261, 1.570796, 2.083853],accel_mss,speed_ms,0,blend_radius_m)
  movel([0.510957, -1.449619, -2.527572, -0.735199, 1.570796, 2.081753],accel_mss,speed_ms,0,blend_radius_m)
  movel([0.508894, -1.449544, -2.527632, -0.735213, 1.570796, 2.079690],accel_mss,speed_ms,0,blend_radius_m)
  movel([0.506952, -1.449051, -2.528029, -0.735309, 1.570796, 2.077748],accel_mss,speed_ms,0,blend_radius_m)
  movel([0.505206, -1.448127, -2.528773, -0.735489, 1.570796, 2.076003],accel_mss,speed_ms,0,blend_radius_m)
  movel([0.503720, -1.446767, -2.529866, -0.735756, 1.570796, 2.074516],accel_mss,speed_ms,0,blend_radius_m)
  movel([0.502541, -1.444964, -2.531310, -0.736115, 1.570796, 2.073337],accel_mss,speed_ms,0,blend_radius_m)
  movel([0.501720, -1.442709, -2.533109, -0.736571, 1.570796, 2.072516],accel_mss,speed_ms,0,blend_radius_m)
  movel([0.501301, -1.439983, -2.535274, -0.737132, 1.570796, 2.072097],accel_mss,speed_ms,0,blend_radius_m)
  movel([0.501294, -1.439855, -2.535375, -0.737159, 1.570796, 2.072091],accel_mss,speed_ms,0,blend_radius_m)
  speed_ms = 0.05
  movel([0.501294, -1.389528, -2.511119, -0.811742, 1.570796, 2.072091],accel_mss,speed_ms,0,blend_radius_m)
  speed_ms = 0.051
  movel([0.501294, -1.380106, -2.506003, -0.826280, 1.570796, 2.072091],accel_mss,speed_ms,0,blend_radius_m)
  movel([0.578727, -1.307215, -2.555223, -0.849950, 1.570796, 2.149524],accel_mss,speed_ms,0,blend_radius_m)
  movel([0.578727, -1.337560, -2.571443, -0.803386, 1.570796, 2.149524],accel_mss,speed_ms,0,blend_radius_m)
  speed_ms = 0.017
  movel([0.578727, -1.370227, -2.586862, -0.755300, 1.570796, 2.149524],accel_mss,speed_ms,0,blend_radius_m)
  speed_ms = 0.051
  movel([0.578353, -1.371010, -2.586322, -0.755057, 1.570796, 2.149149],accel_mss,speed_ms,0,blend_radius_m)
  movel([0.577638, -1.371638, -2.585889, -0.754862, 1.570796, 2.148434],accel_mss,speed_ms,0,blend_radius_m)
  movel([0.576691, -1.372014, -2.585629, -0.754746, 1.570796, 2.147487],accel_mss,speed_ms,0,blend_radius_m)
  movel([0.575826, -1.371951, -2.585672, -0.754765, 1.570796, 2.146622],accel_mss,speed_ms,0,blend_radius_m)
  movel([0.575406, -1.371504, -2.585981, -0.754903, 1.570796, 2.146202],accel_mss,speed_ms,0,blend_radius_m)
  movel([0.573957, -1.369736, -2.587199, -0.755454, 1.570796, 2.144753],accel_mss,speed_ms,0,blend_radius_m)
  movel([0.572628, -1.368361, -2.588144, -0.755884, 1.570796, 2.143424],accel_mss,speed_ms,0,blend_radius_m)
  movel([0.571530, -1.367468, -2.588755, -0.756166, 1.570796, 2.142326],accel_mss,speed_ms,0,blend_radius_m)
  movel([0.570492, -1.366822, -2.589197, -0.756370, 1.570796, 2.141288],accel_mss,speed_ms,0,blend_radius_m)
  movel([0.569467, -1.366363, -2.589511, -0.756515, 1.570796, 2.140263],accel_mss,speed_ms,0,blend_radius_m)
  movel([0.567929, -1.365964, -2.589783, -0.756642, 1.570796, 2.138725],accel_mss,speed_ms,0,blend_radius_m)
  movel([0.566562, -1.365850, -2.589861, -0.756678, 1.570796, 2.137359],accel_mss,speed_ms,0,blend_radius_m)
  movel([0.564121, -1.366028, -2.589739, -0.756621, 1.570796, 2.134917],accel_mss,speed_ms,0,blend_radius_m)
  movel([0.561090, -1.366674, -2.589298, -0.756416, 1.570796, 2.131886],accel_mss,speed_ms,0,blend_radius_m)
  movel([0.557152, -1.367889, -2.588467, -0.756033, 1.570796, 2.127949],accel_mss,speed_ms,0,blend_radius_m)
  movel([0.555681, -1.368393, -2.588122, -0.755874, 1.570796, 2.126477],accel_mss,speed_ms,0,blend_radius_m)
  movel([0.555031, -1.368629, -2.587960, -0.755800, 1.570796, 2.125827],accel_mss,speed_ms,0,blend_radius_m)
  movel([0.554263, -1.368585, -2.587990, -0.755814, 1.570796, 2.125059],accel_mss,speed_ms,0,blend_radius_m)
  movel([0.553752, -1.368122, -2.588308, -0.755960, 1.570796, 2.124548],accel_mss,speed_ms,0,blend_radius_m)
  movel([0.553693, -1.367339, -2.588844, -0.756206, 1.570796, 2.124489],accel_mss,speed_ms,0,blend_radius_m)
  movel([0.553862, -1.366929, -2.589124, -0.756336, 1.570796, 2.124658],accel_mss,speed_ms,0,blend_radius_m)
  movel([0.554502, -1.366195, -2.589626, -0.756569, 1.570796, 2.125298],accel_mss,speed_ms,0,blend_radius_m)
  movel([0.557374, -1.363838, -2.591231, -0.757320, 1.570796, 2.128170],accel_mss,speed_ms,0,blend_radius_m)
  movel([0.559757, -1.361760, -2.592639, -0.757990, 1.570796, 2.130553],accel_mss,speed_ms,0,blend_radius_m)
  movel([0.561359, -1.360221, -2.593678, -0.758490, 1.570796, 2.132155],accel_mss,speed_ms,0,blend_radius_m)
  movel([0.562626, -1.358865, -2.594591, -0.758933, 1.570796, 2.133423],accel_mss,speed_ms,0,blend_radius_m)
  movel([0.563660, -1.357611, -2.595433, -0.759345, 1.570796, 2.134456],accel_mss,speed_ms,0,blend_radius_m)
  movel([0.564917, -1.355772, -2.596664, -0.759953, 1.570796, 2.135713],accel_mss,speed_ms,0,blend_radius_m)
  movel([0.565701, -1.354278, -2.597660, -0.760451, 1.570796, 2.136498],accel_mss,speed_ms,0,blend_radius_m)
  movel([0.566592, -1.351866, -2.599262, -0.761261, 1.570796, 2.137388],accel_mss,speed_ms,0,blend_radius_m)
  movel([0.567189, -1.349060, -2.601115, -0.762214, 1.570796, 2.137985],accel_mss,speed_ms,0,blend_radius_m)
  movel([0.567525, -1.345547, -2.603420, -0.763422, 1.570796, 2.138321],accel_mss,speed_ms,0,blend_radius_m)
  movel([0.567610, -1.343980, -2.604442, -0.763966, 1.570796, 2.138406],accel_mss,speed_ms,0,blend_radius_m)
  movel([0.567758, -1.343384, -2.604830, -0.764175, 1.570796, 2.138555],accel_mss,speed_ms,0,blend_radius_m)
  movel([0.568315, -1.342632, -2.605319, -0.764438, 1.570796, 2.139111],accel_mss,speed_ms,0,blend_radius_m)
  movel([0.569208, -1.342044, -2.605701, -0.764644, 1.570796, 2.140004],accel_mss,speed_ms,0,blend_radius_m)
  movel([0.570214, -1.341817, -2.605848, -0.764724, 1.570796, 2.141010],accel_mss,speed_ms,0,blend_radius_m)
  movel([0.570615, -1.341896, -2.605797, -0.764696, 1.570796, 2.141412],accel_mss,speed_ms,0,blend_radius_m)
  movel([0.571077, -1.342367, -2.605491, -0.764531, 1.570796, 2.141874],accel_mss,speed_ms,0,blend_radius_m)
  movel([0.572582, -1.344184, -2.604309, -0.763895, 1.570796, 2.143378],accel_mss,speed_ms,0,blend_radius_m)
  movel([0.573951, -1.345591, -2.603391, -0.763407, 1.570796, 2.144748],accel_mss,speed_ms,0,blend_radius_m)
  movel([0.575073, -1.346505, -2.602793, -0.763091, 1.570796, 2.145869],accel_mss,speed_ms,0,blend_radius_m)
  movel([0.576133, -1.347166, -2.602359, -0.762863, 1.570796, 2.146929],accel_mss,speed_ms,0,blend_radius_m)
  movel([0.577175, -1.347638, -2.602050, -0.762701, 1.570796, 2.147971],accel_mss,speed_ms,0,blend_radius_m)
  movel([0.578734, -1.348054, -2.601777, -0.762558, 1.570796, 2.149531],accel_mss,speed_ms,0,blend_radius_m)
  movel([0.580125, -1.348174, -2.601698, -0.762517, 1.570796, 2.150921],accel_mss,speed_ms,0,blend_radius_m)
  movel([0.582608, -1.348008, -2.601807, -0.762574, 1.570796, 2.153405],accel_mss,speed_ms,0,blend_radius_m)
  movel([0.585695, -1.347379, -2.602220, -0.762790, 1.570796, 2.156491],accel_mss,speed_ms,0,blend_radius_m)
  movel([0.589724, -1.346187, -2.603001, -0.763201, 1.570796, 2.160520],accel_mss,speed_ms,0,blend_radius_m)
  movel([0.591233, -1.345696, -2.603322, -0.763371, 1.570796, 2.162029],accel_mss,speed_ms,0,blend_radius_m)
  movel([0.591896, -1.345468, -2.603472, -0.763450, 1.570796, 2.162693],accel_mss,speed_ms,0,blend_radius_m)
  movel([0.592664, -1.345537, -2.603426, -0.763426, 1.570796, 2.163461],accel_mss,speed_ms,0,blend_radius_m)
  movel([0.593160, -1.346039, -2.603098, -0.763252, 1.570796, 2.163956],accel_mss,speed_ms,0,blend_radius_m)
  movel([0.593178, -1.346867, -2.602556, -0.762966, 1.570796, 2.163974],accel_mss,speed_ms,0,blend_radius_m)
  movel([0.592988, -1.347292, -2.602277, -0.762820, 1.570796, 2.163785],accel_mss,speed_ms,0,blend_radius_m)
  movel([0.592314, -1.348032, -2.601791, -0.762566, 1.570796, 2.163111],accel_mss,speed_ms,0,blend_radius_m)
  movel([0.589330, -1.350401, -2.600231, -0.761757, 1.570796, 2.160127],accel_mss,speed_ms,0,blend_radius_m)
  movel([0.586877, -1.352480, -2.598855, -0.761054, 1.570796, 2.157673],accel_mss,speed_ms,0,blend_radius_m)
  movel([0.585232, -1.354015, -2.597835, -0.760539, 1.570796, 2.156029],accel_mss,speed_ms,0,blend_radius_m)
  movel([0.583932, -1.355372, -2.596931, -0.760086, 1.570796, 2.154728],accel_mss,speed_ms,0,blend_radius_m)
  movel([0.582872, -1.356620, -2.596096, -0.759672, 1.570796, 2.153669],accel_mss,speed_ms,0,blend_radius_m)
  movel([0.581586, -1.358452, -2.594869, -0.759068, 1.570796, 2.152382],accel_mss,speed_ms,0,blend_radius_m)
  movel([0.580767, -1.359963, -2.593852, -0.758574, 1.570796, 2.151563],accel_mss,speed_ms,0,blend_radius_m)
  movel([0.579860, -1.362325, -2.592257, -0.757807, 1.570796, 2.150656],accel_mss,speed_ms,0,blend_radius_m)
  movel([0.579245, -1.365064, -2.590397, -0.756928, 1.570796, 2.150042],accel_mss,speed_ms,0,blend_radius_m)
  movel([0.578860, -1.368544, -2.588018, -0.755827, 1.570796, 2.149656],accel_mss,speed_ms,0,blend_radius_m)
  movel([0.578727, -1.370227, -2.586862, -0.755300, 1.570796, 2.149524],accel_mss,speed_ms,0,blend_radius_m)
  speed_ms = 0.05
  movel([0.578727, -1.317076, -2.560715, -0.834597, 1.570796, 2.149524],accel_mss,speed_ms,0,blend_radius_m)
  speed_ms = 0.051
  movel([0.578727, -1.307215, -2.555223, -0.849950, 1.570796, 2.149524],accel_mss,speed_ms,0,blend_radius_m)
  movel([0.341909, -1.348942, -2.527901, -0.835546, 1.570796, 1.912706],accel_mss,speed_ms,0,blend_radius_m)
  movel([0.341909, -1.378495, -2.543467, -0.790428, 1.570796, 1.912706],accel_mss,speed_ms,0,blend_radius_m)
  speed_ms = 0.017
  movel([0.341909, -1.410141, -2.558229, -0.744019, 1.570796, 1.912706],accel_mss,speed_ms,0,blend_radius_m)
  speed_ms = 0.051
  movel([0.341733, -1.410741, -2.557781, -0.743867, 1.570796, 1.912529],accel_mss,speed_ms,0,blend_radius_m)
  movel([0.341182, -1.411271, -2.557385, -0.743734, 1.570796, 1.911979],accel_mss,speed_ms,0,blend_radius_m)
  movel([0.340404, -1.411569, -2.557161, -0.743659, 1.570796, 1.911200],accel_mss,speed_ms,0,blend_radius_m)
  movel([0.340058, -1.411553, -2.557173, -0.743663, 1.570796, 1.910855],accel_mss,speed_ms,0,blend_radius_m)
  movel([0.339733, -1.411364, -2.557315, -0.743710, 1.570796, 1.910529],accel_mss,speed_ms,0,blend_radius_m)
  movel([0.338240, -1.410318, -2.558097, -0.743974, 1.570796, 1.909036],accel_mss,speed_ms,0,blend_radius_m)
  movel([0.336366, -1.409558, -2.558665, -0.744167, 1.570796, 1.907163],accel_mss,speed_ms,0,blend_radius_m)
  movel([0.334413, -1.409267, -2.558881, -0.744241, 1.570796, 1.905209],accel_mss,speed_ms,0,blend_radius_m)
  movel([0.332363, -1.409394, -2.558787, -0.744208, 1.570796, 1.903160],accel_mss,speed_ms,0,blend_radius_m)
  movel([0.330181, -1.409911, -2.558401, -0.744077, 1.570796, 1.900977],accel_mss,speed_ms,0,blend_radius_m)
  movel([0.327818, -1.410814, -2.557726, -0.743849, 1.570796, 1.898614],accel_mss,speed_ms,0,blend_radius_m)
  movel([0.325137, -1.412092, -2.556769, -0.743527, 1.570796, 1.895933],accel_mss,speed_ms,0,blend_radius_m)
  movel([0.323918, -1.412588, -2.556397, -0.743403, 1.570796, 1.894714],accel_mss,speed_ms,0,blend_radius_m)
  movel([0.323545, -1.412630, -2.556366, -0.743393, 1.570796, 1.894341],accel_mss,speed_ms,0,blend_radius_m)
  movel([0.323353, -1.412549, -2.556427, -0.743413, 1.570796, 1.894150],accel_mss,speed_ms,0,blend_radius_m)
  movel([0.323276, -1.412068, -2.556788, -0.743534, 1.570796, 1.894072],accel_mss,speed_ms,0,blend_radius_m)
  movel([0.323548, -1.411192, -2.557444, -0.743753, 1.570796, 1.894344],accel_mss,speed_ms,0,blend_radius_m)
  movel([0.326783, -1.407562, -2.560150, -0.744677, 1.570796, 1.897580],accel_mss,speed_ms,0,blend_radius_m)
  movel([0.327727, -1.406298, -2.561088, -0.745003, 1.570796, 1.898523],accel_mss,speed_ms,0,blend_radius_m)
  movel([0.328413, -1.405209, -2.561894, -0.745286, 1.570796, 1.899210],accel_mss,speed_ms,0,blend_radius_m)
  movel([0.329132, -1.403689, -2.563016, -0.745684, 1.570796, 1.899929],accel_mss,speed_ms,0,blend_radius_m)
  movel([0.329417, -1.402715, -2.563734, -0.745940, 1.570796, 1.900214],accel_mss,speed_ms,0,blend_radius_m)
  movel([0.329610, -1.400922, -2.565050, -0.746417, 1.570796, 1.900406],accel_mss,speed_ms,0,blend_radius_m)
  movel([0.329403, -1.398862, -2.566557, -0.746970, 1.570796, 1.900199],accel_mss,speed_ms,0,blend_radius_m)
  movel([0.328847, -1.396525, -2.568259, -0.747605, 1.570796, 1.899643],accel_mss,speed_ms,0,blend_radius_m)
  movel([0.329185, -1.395686, -2.568868, -0.747835, 1.570796, 1.899981],accel_mss,speed_ms,0,blend_radius_m)
  movel([0.329453, -1.395281, -2.569162, -0.747946, 1.570796, 1.900249],accel_mss,speed_ms,0,blend_radius_m)
  movel([0.329701, -1.395069, -2.569315, -0.748005, 1.570796, 1.900498],accel_mss,speed_ms,0,blend_radius_m)
  movel([0.330225, -1.394952, -2.569400, -0.748037, 1.570796, 1.901022],accel_mss,speed_ms,0,blend_radius_m)
  movel([0.331042, -1.395216, -2.569209, -0.747964, 1.570796, 1.901838],accel_mss,speed_ms,0,blend_radius_m)
  movel([0.333110, -1.396285, -2.568434, -0.747671, 1.570796, 1.903907],accel_mss,speed_ms,0,blend_radius_m)
  movel([0.334370, -1.396763, -2.568086, -0.747540, 1.570796, 1.905167],accel_mss,speed_ms,0,blend_radius_m)
  movel([0.335488, -1.397033, -2.567890, -0.747466, 1.570796, 1.906284],accel_mss,speed_ms,0,blend_radius_m)
  movel([0.336585, -1.397163, -2.567795, -0.747431, 1.570796, 1.907382],accel_mss,speed_ms,0,blend_radius_m)
  movel([0.337693, -1.397169, -2.567791, -0.747429, 1.570796, 1.908489],accel_mss,speed_ms,0,blend_radius_m)
  movel([0.338826, -1.397058, -2.567871, -0.747459, 1.570796, 1.909623],accel_mss,speed_ms,0,blend_radius_m)
  movel([0.341268, -1.396472, -2.568298, -0.747619, 1.570796, 1.912064],accel_mss,speed_ms,0,blend_radius_m)
  movel([0.343929, -1.395382, -2.569089, -0.747918, 1.570796, 1.914726],accel_mss,speed_ms,0,blend_radius_m)
  movel([0.346252, -1.394117, -2.570005, -0.748268, 1.570796, 1.917048],accel_mss,speed_ms,0,blend_radius_m)
  movel([0.346742, -1.393871, -2.570182, -0.748336, 1.570796, 1.917538],accel_mss,speed_ms,0,blend_radius_m)
  movel([0.347389, -1.393839, -2.570205, -0.748345, 1.570796, 1.918185],accel_mss,speed_ms,0,blend_radius_m)
  movel([0.347817, -1.394202, -2.569943, -0.748244, 1.570796, 1.918613],accel_mss,speed_ms,0,blend_radius_m)
  movel([0.347796, -1.394865, -2.569463, -0.748061, 1.570796, 1.918593],accel_mss,speed_ms,0,blend_radius_m)
  movel([0.347278, -1.395523, -2.568986, -0.747880, 1.570796, 1.918074],accel_mss,speed_ms,0,blend_radius_m)
  movel([0.345358, -1.397439, -2.567595, -0.747356, 1.570796, 1.916154],accel_mss,speed_ms,0,blend_radius_m)
  movel([0.343566, -1.399686, -2.565955, -0.746748, 1.570796, 1.914363],accel_mss,speed_ms,0,blend_radius_m)
  movel([0.342312, -1.401850, -2.564369, -0.746170, 1.570796, 1.913108],accel_mss,speed_ms,0,blend_radius_m)
  movel([0.341536, -1.403970, -2.562809, -0.745610, 1.570796, 1.912332],accel_mss,speed_ms,0,blend_radius_m)
  movel([0.341217, -1.406083, -2.561247, -0.745059, 1.570796, 1.912013],accel_mss,speed_ms,0,blend_radius_m)
  movel([0.341362, -1.408224, -2.559658, -0.744507, 1.570796, 1.912159],accel_mss,speed_ms,0,blend_radius_m)
  movel([0.341909, -1.410141, -2.558229, -0.744019, 1.570796, 1.912706],accel_mss,speed_ms,0,blend_radius_m)
  speed_ms = 0.05
  movel([0.341909, -1.348942, -2.527901, -0.835546, 1.570796, 1.912706],accel_mss,speed_ms,0,blend_radius_m)
  movel([0.341909, -1.295920, -2.494548, -0.921922, 1.570796, 1.912706],accel_mss,speed_ms,0,blend_radius_m)
  #M_RunCode5
  #M_RunCode30
  # End of main program
end

Machining1()
